Fanuc KAREL source: KO00129.KL

PROGRAM KO00129
%NOLOCKGROUP
VAR
  R: REAL
  CFG: CONFIG
  OUT: XYZWPR
  N: INTEGER
BEGIN
  N = 1
  R = 2.0
  CFG.CFG_FLIP = TRUE
  OUT = POS(N, R, R, R, R, R, CFG)
END KO00129
